TYPE ST_Blinker_1 :
STRUCT	
	Q0					:BOOL; 						(* Divider output / 2 *)
	Q1					:BOOL; 						(* Divider output / 4 *)
	Q2					:BOOL; 						(* Divider output / 8 *)
	Q3					:BOOL; 						(* Divider output / 16 *)
	Q4					:BOOL; 						(* Divider output / 32 *)
	Q5					:BOOL; 						(* Divider output / 64 *)
	Q6					:BOOL; 						(* Divider output / 128 *)
	Q7					:BOOL; 						(* Divider output / 256 *)
END_STRUCT
END_TYPE

(* stored: Version 1.1.0.1, ProductVersion 3.1.4024.15
   DUT ST_Blinker_1: Id {04db8fb6-9352-4188-b0dd-9cc073e15e52} *)
